(* PLC project g_burner_purge_self_clearing, Anonymous Benchmark Suite 1.0 *)
(* stored: creationDateTime 2026-08-28T00:00:00 *)

PROGRAM g_burner_purge_self_clearing
  VAR_INPUT
    CallForHeat : BOOL;
    PurgeDone : BOOL;
    FlameProven : BOOL;
    FlameFail : BOOL;
    ResetBtn : BOOL;
  END_VAR
  VAR_OUTPUT
    Fan : BOOL;
    Lockout : BOOL;
    Pilot : BOOL;
    MainValve : BOOL;
  END_VAR

(* LD diagram, written out as Structured Text *)
Fan := CallForHeat;
Lockout := FlameFail AND NOT ResetBtn;
Pilot := CallForHeat AND PurgeDone AND NOT Lockout;
MainValve := CallForHeat AND PurgeDone AND FlameProven AND NOT Lockout;
END_PROGRAM

CONFIGURATION Config0
  RESOURCE Res0 ON PLC
    TASK tcyclic(INTERVAL := T#10ms, PRIORITY := 0);
    PROGRAM inst0 WITH tcyclic : g_burner_purge_self_clearing;
  END_RESOURCE
END_CONFIGURATION
